Fanuc KAREL source: kc00026.KL

-- PROVISIONAL review KL for V1013-1; original PC SHA256 85842cd8e93cfcf412d3fdb6acdc619512d3c43c29c474afbc2197cdf2e6b830
-- Incomplete behavior may be omitted. Consult companion uncertainty JSON. Do not deploy.
PROGRAM KC00026
%NOLOCKGROUP
BEGIN
  -- UNRESOLVED_PC offsets 5-45; opcodes 27,22,22,22,22,22,22,31
  -- UNRESOLVED_PC offsets 50-54; opcodes 7F
END KC00026
